// CFC twin of T_SafeAnd_Tests: the same tests drawn as CFC diagrams, the way a TwinSAFE project is authored.
    FUNCTION_BLOCK T_SafeAnd_Tests_CFC EXTENDS T_SafeCfcTestSuite
    VAR
    // Test_AllConnectedInputsTrueGivesRun
    group_1 : T_SafeGroup;
    fb_1 : T_SafeAnd(group := group_1);
    // Test_OneInputFalseGivesSafe
    group_2 : T_SafeGroup;
    fb_2 : T_SafeAnd(group := group_2);
    // Test_UnconnectedInputsIgnoredAndMakeContactNegated
    group_3 : T_SafeGroup;
    fb_3 : T_SafeAnd(group := group_3) := (Parameters := (In2MakeContact := TRUE));
    // Test_StoppedGivesNoOutput
    group_4 : T_SafeGroup;
    fb_4 : T_SafeAnd(group := group_4);
END_VAR

Test_AllConnectedInputsTrueGivesRun();
Test_OneInputFalseGivesSafe();
Test_UnconnectedInputsIgnoredAndMakeContactNegated();
Test_StoppedGivesNoOutput();

METHOD PRIVATE Test_AllConnectedInputsTrueGivesRun
// note: this text did not pass the execution check against the stored diagram
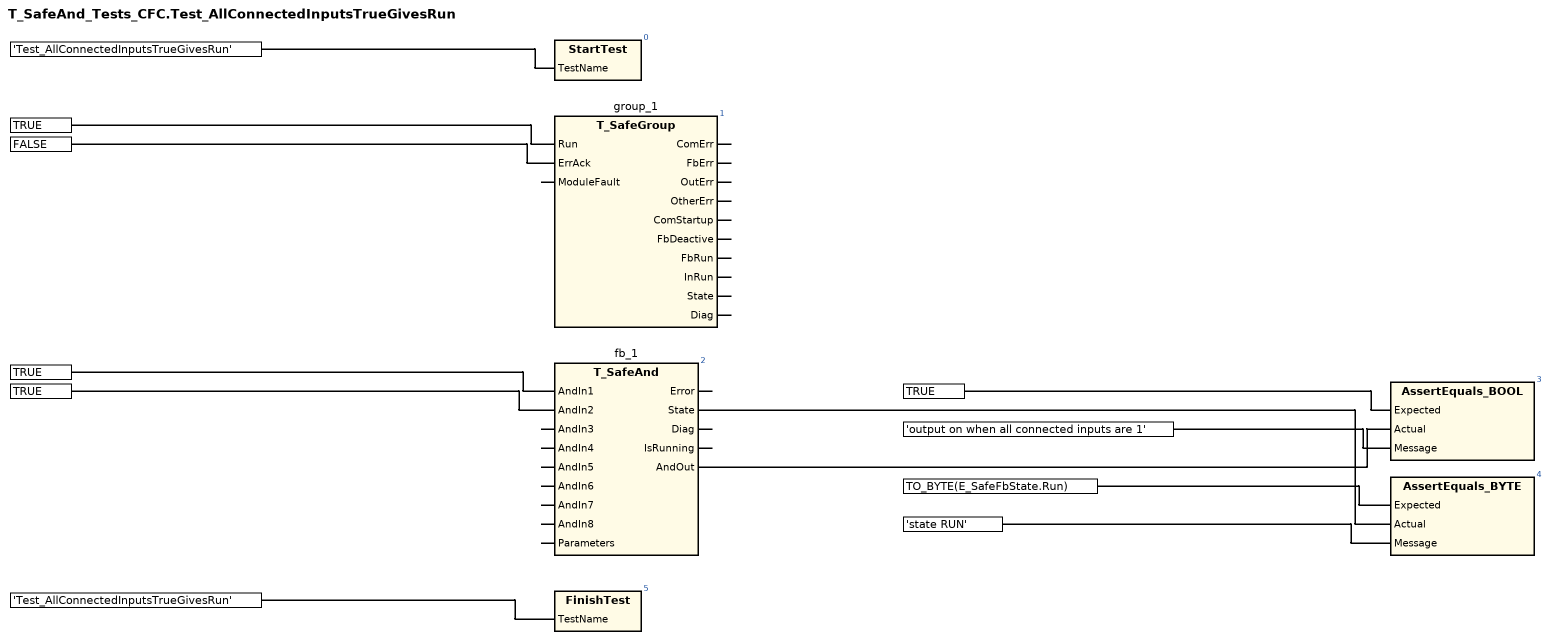
StartTest(TestName := 'Test_AllConnectedInputsTrueGivesRun');
group_1(Run := TRUE, ErrAck := FALSE); // T_SafeGroup
fb_1(AndIn1 := TRUE, AndIn2 := TRUE); // T_SafeAnd
AssertEquals_BOOL(Expected := TRUE, Actual := fb_1.AndOut, Message := 'output on when all connected inputs are 1');
AssertEquals_BYTE(Expected := TO_BYTE(E_SafeFbState.Run), Actual := fb_1.State, Message := 'state RUN');
FinishTest(TestName := 'Test_AllConnectedInputsTrueGivesRun');
END_METHOD

METHOD PRIVATE Test_OneInputFalseGivesSafe
// note: this text did not pass the execution check against the stored diagram
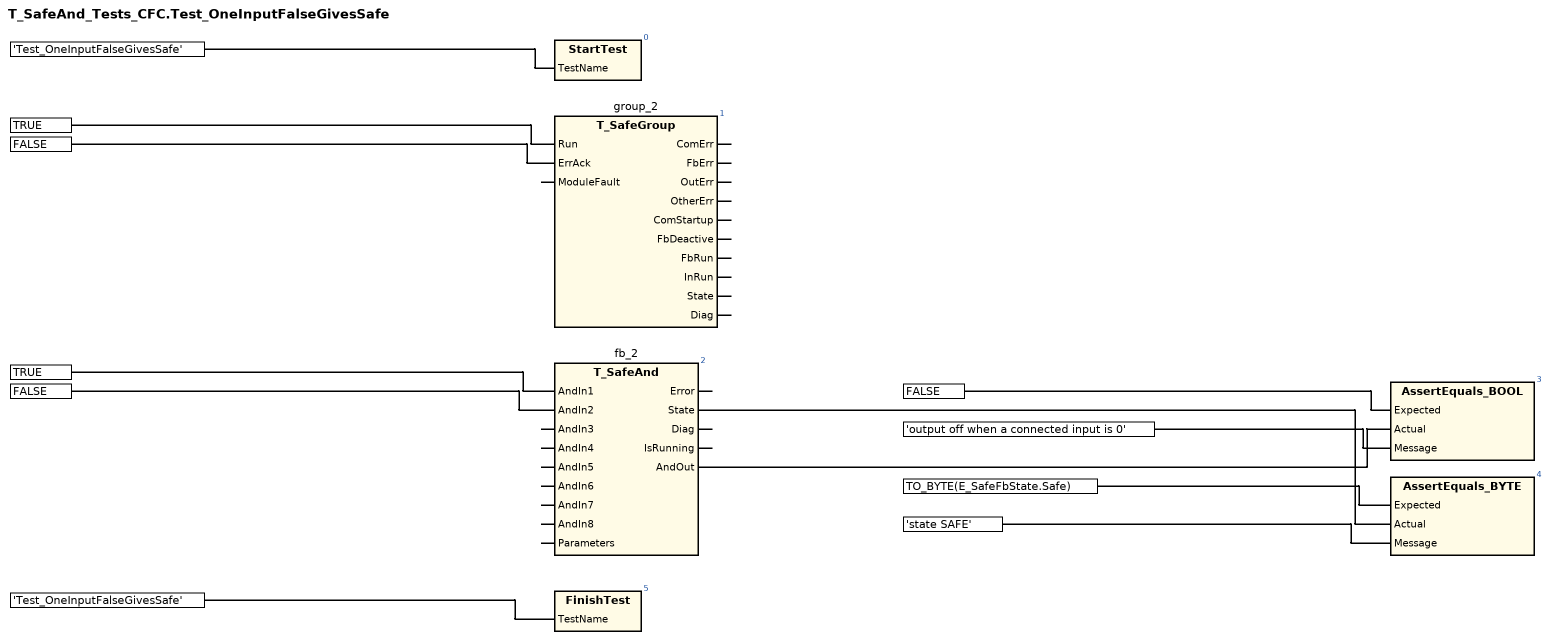
StartTest(TestName := 'Test_OneInputFalseGivesSafe');
group_2(Run := TRUE, ErrAck := FALSE); // T_SafeGroup
fb_2(AndIn1 := TRUE, AndIn2 := FALSE); // T_SafeAnd
AssertEquals_BOOL(Expected := FALSE, Actual := fb_2.AndOut, Message := 'output off when a connected input is 0');
AssertEquals_BYTE(Expected := TO_BYTE(E_SafeFbState.Safe), Actual := fb_2.State, Message := 'state SAFE');
FinishTest(TestName := 'Test_OneInputFalseGivesSafe');
END_METHOD

METHOD PRIVATE Test_UnconnectedInputsIgnoredAndMakeContactNegated
// note: this text did not pass the execution check against the stored diagram
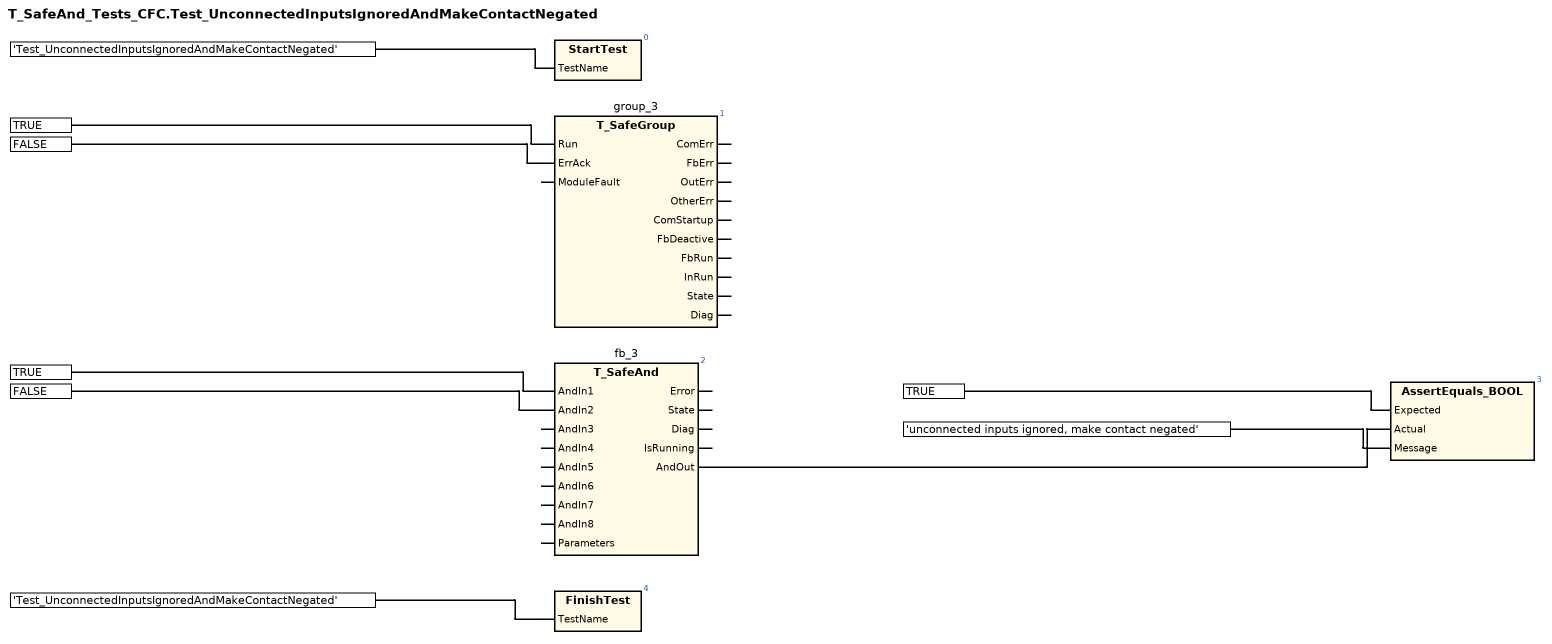
StartTest(TestName := 'Test_UnconnectedInputsIgnoredAndMakeContactNegated');
group_3(Run := TRUE, ErrAck := FALSE); // T_SafeGroup
fb_3(AndIn1 := TRUE, AndIn2 := FALSE); // T_SafeAnd
AssertEquals_BOOL(Expected := TRUE, Actual := fb_3.AndOut, Message := 'unconnected inputs ignored, make contact negated');
FinishTest(TestName := 'Test_UnconnectedInputsIgnoredAndMakeContactNegated');
END_METHOD

METHOD PRIVATE Test_StoppedGivesNoOutput
// note: this text did not pass the execution check against the stored diagram
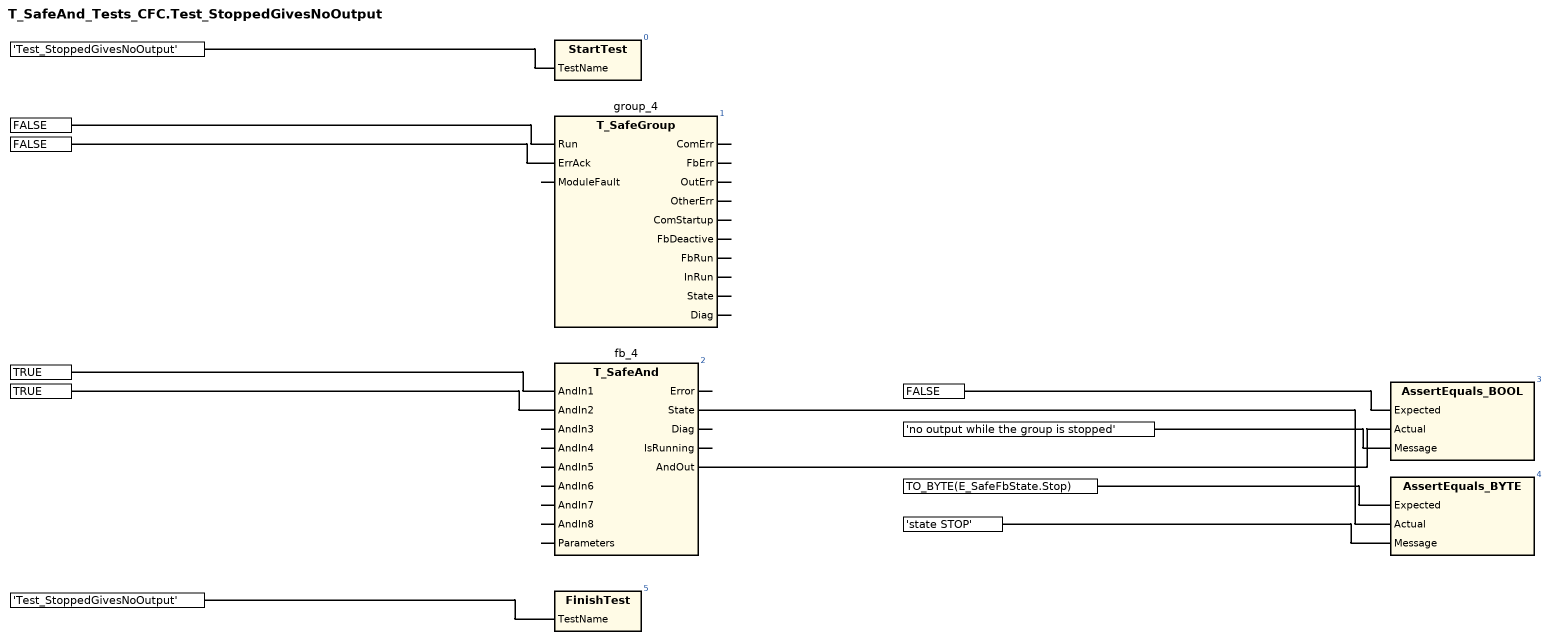
StartTest(TestName := 'Test_StoppedGivesNoOutput');
group_4(Run := FALSE, ErrAck := FALSE); // T_SafeGroup
fb_4(AndIn1 := TRUE, AndIn2 := TRUE); // T_SafeAnd
AssertEquals_BOOL(Expected := FALSE, Actual := fb_4.AndOut, Message := 'no output while the group is stopped');
AssertEquals_BYTE(Expected := TO_BYTE(E_SafeFbState.Stop), Actual := fb_4.State, Message := 'state STOP');
FinishTest(TestName := 'Test_StoppedGivesNoOutput');
END_METHOD

END_FUNCTION_BLOCK

(* stored: Version 1.1.0.1, ProductVersion 3.1.4026.22
   POU T_SafeAnd_Tests_CFC: Id {0f19d271-aa04-5ab9-846c-ea140fc85df3}, SpecialFunc None
   Method Test_AllConnectedInputsTrueGivesRun: Id {6a2bf4ac-c7e2-50c2-b146-141d4bd6a23b}
   Method Test_OneInputFalseGivesSafe: Id {950ddba0-71ee-519d-8de9-b9f218fc9bb2}
   Method Test_UnconnectedInputsIgnoredAndMakeContactNegated: Id {c553b8b0-7ebc-5c5c-86ca-f51d61d685c6}
   Method Test_StoppedGivesNoOutput: Id {076bb0a4-0866-5960-9e6f-8189019340c6} *)
